Staubli VAL3: safePointCheck.pgx

public program safePointCheck()
  local bool l_bResult
  local bool l_bErr
  local num l_i
begin
  for l_i = 0 to size(safeTemp:sSPoint)-1
    call computeSPoint(l_i,l_bResult)
    //O_safePoint[l_i]=(l_bResult==true)
    call io:setDigOutput(O_safePoint[l_i],l_bResult,l_bErr)
  endFor
end
